Fanuc KAREL source: kb00156.KL

-- PROVISIONAL review KL for V1013-1; original PC SHA256 509b12f32e19a9ec0fe0c306cac354af437dbae2b4f70c92c365a1a61374f2b3
-- Incomplete behavior may be omitted. Consult companion uncertainty JSON. Do not deploy.
PROGRAM KB00156
%NOLOCKGROUP
BEGIN
  -- UNRESOLVED_PC offsets 5-14; opcodes 3F,75
  -- UNRESOLVED_PC offsets 19-26; opcodes 9D,23
  -- UNRESOLVED_PC offsets 31-49; opcodes 27,22,2A,22,31
  -- UNRESOLVED_PC offsets 54-58; opcodes 7F
END KB00156
